(* IEC 61131-3 sources: STAR-PLC-Agent/results/raw/codex_matrix_resume_20261114/codex_terra/SELF001/formal/attempt_0001, 1 file *)

(* ---- candidate.st ---- *)
FUNCTION_BLOCK FB_Task
VAR_INPUT
    Start : BOOL;
    Stop : BOOL;
    GuardClosed : BOOL;
END_VAR
VAR_OUTPUT
    Run : BOOL := FALSE;
END_VAR

IF Stop OR NOT GuardClosed THEN
    Run := FALSE;
ELSIF Start THEN
    Run := TRUE;
END_IF;
END_FUNCTION_BLOCK
